(*
	Owned collection of OTLP key-value attributes used across telemetry domains.
*)
{attribute 'enable_dynamic_creation'}
FUNCTION_BLOCK FB_Attributes
VAR
	_head: POINTER TO ST_LinkedListNode;
	_tail: POINTER TO ST_LinkedListNode;
	_cursor: POINTER TO ST_LinkedListNode;
END_VAR
VAR_OUTPUT
	count: UDINT;
	maxCount: UDINT;
	droppedCount: UDINT;
END_VAR

(* The enforced bound: maxCount, held to MAX_LOOP_COUNT so free always reaches the end. *)
METHOD _capacity : UDINT
_capacity := MIN(THIS^.maxCount, TcOtlp_GVL.MAX_LOOP_COUNT);
END_METHOD

(* The node holding the attribute named key, or 0 when there is none. Does not move the next cursor. *)
METHOD _findNode : POINTER TO ST_LinkedListNode
VAR_INPUT
	key: T_MaxString;
END_VAR
VAR
	_idx: UDINT;
	_node: POINTER TO ST_LinkedListNode;
	_pKv: POINTER TO FB_KeyValue;
END_VAR
_findNode := 0;

_node := THIS^._head;
FOR _idx := 0 TO TcOtlp_GVL.MAX_LOOP_COUNT DO
	IF _node = 0 THEN
		RETURN;
	END_IF
	_pKv := _node^.val;
	IF _pKv <> 0 AND_THEN _pKv^.pKey <> 0 AND_THEN _pKv^.pKey^ = key THEN
		_findNode := _node;
		RETURN;
	END_IF
	_node := _node^.nxt;
END_FOR
END_METHOD

METHOD _mapValueFactoryFailure : E_AttributesFailureReason
VAR_INPUT
	failureReason: E_ValueFactoryFailureReason;
END_VAR
CASE failureReason OF
	E_ValueFactoryFailureReason.SOURCE_POINTER_NULL:
		_mapValueFactoryFailure := E_AttributesFailureReason.KV_VALUE_POINTER_NULL;
	E_ValueFactoryFailureReason.KEY_POINTER_NULL:
		_mapValueFactoryFailure := E_AttributesFailureReason.KV_KEY_POINTER_NULL;
	E_ValueFactoryFailureReason.VALUE_POINTER_NULL:
		_mapValueFactoryFailure := E_AttributesFailureReason.KV_VALUE_POINTER_NULL;
	E_ValueFactoryFailureReason.UNSUPPORTED_VALUE_TYPE:
		_mapValueFactoryFailure := E_AttributesFailureReason.KV_VALUE_TYPE_UNSUPPORTED;
	E_ValueFactoryFailureReason.MEMORY_ALLOCATION_FAILURE:
		_mapValueFactoryFailure := E_AttributesFailureReason.MEMORY_ALLOCATION_FAILURE;
	ELSE
		_mapValueFactoryFailure := E_AttributesFailureReason.KV_VALUE_INVALID;
END_CASE
END_METHOD

(*
	Adds a copy of src's attribute named key, stored under destKey, or under key when destKey is
	empty. An attribute already held under that name is replaced, as with setAttribute. src is
	left unchanged and may be this collection, so an attribute can be copied to a new name in place.
*)
METHOD copyAttribute : BOOL
VAR_IN_OUT
	src: FB_Attributes;
END_VAR
VAR_INPUT
	key: T_MaxString;
	destKey: T_MaxString := '';
END_VAR
VAR_OUTPUT
	failureReason: E_AttributesFailureReason;
END_VAR
VAR
	_pSrc: POINTER TO FB_KeyValue;
	_pDest: POINTER TO FB_KeyValue;
	_factoryFailureReason: E_ValueFactoryFailureReason;
END_VAR
copyAttribute := FALSE;
failureReason := E_AttributesFailureReason.NA;

_pSrc := src.getAttribute(key);
IF _pSrc = 0 THEN
	failureReason := E_AttributesFailureReason.KEY_NOT_FOUND;
	RETURN;
END_IF

IF destKey = '' THEN
	destKey := key;
END_IF

IF NOT ValueFactory.createKeyValue(
	pDest:=_pDest,
	pKey:=ADR(destKey),
	pVal:=_pSrc^.pVal,
	failureReason=>_factoryFailureReason
) THEN
	failureReason := THIS^._mapValueFactoryFailure(_factoryFailureReason);
	RETURN;
END_IF

copyAttribute := THIS^.setAttribute(pValue:=_pDest, failureReason=>failureReason);
// setAttribute only takes ownership on success; release a rejected value
IF _pDest <> 0 THEN
	_pDest^.delete(pSelf:=_pDest);
END_IF
END_METHOD

(*
	Adds a copy of every attribute in src, and carries src's droppedCount over, so the copy
	reports the same loss as the original.
*)
METHOD copyFrom : BOOL
VAR_IN_OUT
	src: FB_Attributes;
END_VAR
VAR_OUTPUT
	failureReason: E_AttributesFailureReason;
END_VAR
VAR
	_idx: UDINT;
	_pSrc: POINTER TO FB_KeyValue;
	_pDest: POINTER TO FB_KeyValue;
	_factoryFailureReason: E_ValueFactoryFailureReason;
END_VAR
copyFrom := FALSE;
failureReason := E_AttributesFailureReason.NA;

THIS^.droppedCount := THIS^.droppedCount + src.droppedCount;
src.reset();
FOR _idx := 0 TO TcOtlp_GVL.MAX_LOOP_COUNT DO
	_pSrc := src.next();
	IF _pSrc = 0 THEN
		copyFrom := failureReason = E_AttributesFailureReason.NA;
		RETURN;
	END_IF
	IF NOT ValueFactory.cloneKeyValue(pDest:=_pDest, pSrc:=_pSrc, failureReason=>_factoryFailureReason) THEN
		failureReason := THIS^._mapValueFactoryFailure(_factoryFailureReason);
		RETURN;
	END_IF
	IF NOT THIS^.setAttribute(pValue:=_pDest, failureReason=>failureReason) THEN
		IF _pDest <> 0 THEN
			_pDest^.delete(pSelf:=_pDest);
		END_IF
		RETURN;
	END_IF
END_FOR

copyFrom := failureReason = E_AttributesFailureReason.NA;
END_METHOD

METHOD FB_Exit : BOOL
VAR_INPUT
	bInCopyCode: BOOL;
END_VAR
IF NOT bInCopyCode THEN
	THIS^.free();
END_IF
END_METHOD

//FB_Init is always available implicitly and it is used primarily for initialization.
//The return value is not evaluated. For a specific influence, you can also declare the
//methods explicitly and provide additional code there with the standard initialization
//code. You can evaluate the return value.
METHOD FB_Init: BOOL
VAR_INPUT
    bInitRetains: BOOL; // TRUE: the retain variables are initialized (reset warm / reset cold)
    bInCopyCode: BOOL;  // TRUE: the instance will be copied to the copy code afterward (online change) 
	maxCount: UDINT := 20;  
END_VAR
THIS^.maxCount := maxCount;
END_METHOD

(*
	Releases every owned attribute. setAttribute holds count to MAX_LOOP_COUNT, so the loop
	always reaches the end, even if maxCount is lowered after attributes were added. If it ever
	stops early, the unreleased nodes stay in the collection and free returns FALSE, so a later
	call can finish the job.
*)
METHOD free : BOOL
VAR
	_idx: UDINT;
	_node: POINTER TO ST_LinkedListNode;
	_kv: POINTER TO FB_KeyValue;
END_VAR
FOR _idx := 0 TO TcOtlp_GVL.MAX_LOOP_COUNT DO
	IF THIS^._head = 0 THEN
		EXIT;
	END_IF

	_node := THIS^._head;
	THIS^._head := _node^.nxt;
	IF _node^.val <> 0 THEN
		_kv := _node^.val;
		_node^.val := 0;
		_kv^.delete(pSelf:=_kv);
	END_IF
	__DELETE(_node);
	_node := 0;
	IF THIS^.count > 0 THEN
		THIS^.count := THIS^.count - 1;
	END_IF
END_FOR

IF THIS^._head = 0 THEN
	THIS^._tail := 0;
	THIS^.count := 0;
END_IF
THIS^._cursor := THIS^._head;
free := THIS^._head = 0;
END_METHOD

(*
	Returns the attribute named key, or 0 when there is none. The collection keeps ownership: the
	pointer is borrowed and stays valid only until that attribute is replaced or the collection is
	freed. Does not move the next cursor.
*)
METHOD getAttribute : POINTER TO FB_KeyValue
VAR_INPUT
	key: T_MaxString;
END_VAR
VAR
	_node: POINTER TO ST_LinkedListNode;
END_VAR
getAttribute := 0;

_node := THIS^._findNode(key);
IF _node <> 0 THEN
	getAttribute := _node^.val;
END_IF
END_METHOD

METHOD next : POINTER TO FB_KeyValue
next := 0;

IF THIS^._cursor <> 0 THEN
	next := THIS^._cursor^.val;
	THIS^._cursor := THIS^._cursor^.nxt;
END_IF
END_METHOD

METHOD reset
THIS^._cursor := THIS^._head;
END_METHOD

METHOD setAttribute : BOOL
VAR_IN_OUT
	pValue: POINTER TO FB_KeyValue;
END_VAR
VAR_OUTPUT
	failureReason: E_AttributesFailureReason;
END_VAR
VAR
	_node: POINTER TO ST_LinkedListNode;
	_pVal: POINTER TO FB_KeyValue;
END_VAR
setAttribute := FALSE;
failureReason := E_AttributesFailureReason.NA;

IF pValue = 0 THEN
	failureReason := E_AttributesFailureReason.KV_POINTER_NULL;
	RETURN;
END_IF

IF pValue^.pKey = 0 THEN
	failureReason := E_AttributesFailureReason.KV_KEY_POINTER_NULL;
	RETURN;
END_IF

IF pValue^.pVal = 0 THEN
	failureReason := E_AttributesFailureReason.KV_VALUE_POINTER_NULL;
	RETURN;
END_IF

// replace the value if the key already exists
_node := THIS^._findNode(pValue^.pKey^);
IF _node <> 0 THEN
	_pVal := _node^.val;
	_pVal^.delete(pSelf:=_pVal);
	_node^.val := pValue;
	setAttribute := failureReason = E_AttributesFailureReason.NA;
	pValue := 0;
	RETURN;
END_IF

IF THIS^.count >= THIS^._capacity() THEN
	failureReason := E_AttributesFailureReason.ATTRIBUTE_COUNT_LIMIT_REACHED;
	THIS^.droppedCount := THIS^.droppedCount + 1;
	RETURN;
END_IF

// if it doesn't exist append the key-value pair
_node := __NEW(ST_LinkedListNode);
IF _node = 0 THEN
	failureReason := E_AttributesFailureReason.MEMORY_ALLOCATION_FAILURE;
	RETURN;
END_IF

_node^.val := pValue;
_node^.nxt := 0;

IF THIS^._tail = 0 THEN
	THIS^._head := _node;
	THIS^._cursor := _node;
ELSE
	THIS^._tail^.nxt := _node;
END_IF

THIS^._tail := _node;
THIS^.count := THIS^.count + 1;

// Ownership transfers only after the value has been linked successfully.
pValue := 0;
setAttribute := failureReason = E_AttributesFailureReason.NA;
END_METHOD

METHOD setNumberAttribute : BOOL
VAR_INPUT
	key: T_MaxString;
	value: ANY_NUM;
END_VAR
VAR_OUTPUT
	failureReason: E_AttributesFailureReason;
END_VAR
VAR
	_pKv: POINTER TO FB_KeyValue;
	_pNum: POINTER TO FB_Number;
	_factoryFailureReason: E_ValueFactoryFailureReason;
END_VAR
setNumberAttribute := FALSE;
failureReason := E_AttributesFailureReason.NA;

IF NOT ValueFactory.createNumber_AnyType(
	pDest:=_pNum,
	value:=value,
	failureReason=>_factoryFailureReason
) THEN
	failureReason := THIS^._mapValueFactoryFailure(_factoryFailureReason);
	RETURN;
END_IF

IF NOT ValueFactory.createKeyValue(
	pDest:=_pKv,
	pKey:=ADR(key),
	pVal:=_pNum,
	failureReason=>_factoryFailureReason
) THEN
	failureReason := THIS^._mapValueFactoryFailure(_factoryFailureReason);
	_pNum^.delete(pSelf:=_pNum);
	RETURN;
END_IF
_pNum^.delete(pSelf:=_pNum);  // clean up the _pNum as its cloned in createKeyValue

setNumberAttribute := THIS^.setAttribute(pValue:=_pKv, failureReason=>failureReason);
// setAttribute only takes ownership on success; release a rejected value
IF _pKv <> 0 THEN
	_pKv^.delete(pSelf:=_pKv);
END_IF
END_METHOD

METHOD setNumberAttribute_AnyType : BOOL
VAR_INPUT
	key: T_MaxString;
	value: AnyType;
END_VAR
VAR_OUTPUT
	failureReason: E_AttributesFailureReason;
END_VAR
VAR
	_pKv: POINTER TO FB_KeyValue;
	_pNum: POINTER TO FB_Number;
	_factoryFailureReason: E_ValueFactoryFailureReason;
END_VAR
setNumberAttribute_AnyType := FALSE;
failureReason := E_AttributesFailureReason.NA;

IF NOT ValueFactory.createNumber_AnyType(
	pDest:=_pNum,
	value:=value,
	failureReason=>_factoryFailureReason
) THEN
	failureReason := THIS^._mapValueFactoryFailure(_factoryFailureReason);
	RETURN;
END_IF

IF NOT ValueFactory.createKeyValue(
	pDest:=_pKv,
	pKey:=ADR(key),
	pVal:=_pNum,
	failureReason=>_factoryFailureReason
) THEN
	failureReason := THIS^._mapValueFactoryFailure(_factoryFailureReason);
	_pNum^.delete(pSelf:=_pNum);
	RETURN;
END_IF
_pNum^.delete(pSelf:=_pNum);  // clean up the _pNum as its cloned in createKeyValue

setNumberAttribute_AnyType := THIS^.setAttribute(pValue:=_pKv, failureReason=>failureReason);
// setAttribute only takes ownership on success; release a rejected value
IF _pKv <> 0 THEN
	_pKv^.delete(pSelf:=_pKv);
END_IF
END_METHOD

METHOD setStringAttribute : BOOL
VAR_INPUT
	key: T_MaxString;
	value: T_MaxString;
END_VAR
VAR_OUTPUT
	failureReason: E_AttributesFailureReason;
END_VAR
VAR
	_pKv: POINTER TO FB_KeyValue;
	_pStr: POINTER TO FB_String;
	_factoryFailureReason: E_ValueFactoryFailureReason;
END_VAR
setStringAttribute := FALSE;
failureReason := E_AttributesFailureReason.NA;

IF NOT ValueFactory.createString(
	pDest:=_pStr,
	pString:=ADR(value),
	failureReason=>_factoryFailureReason
) THEN
	failureReason := THIS^._mapValueFactoryFailure(_factoryFailureReason);
	RETURN;
END_IF

IF NOT ValueFactory.createKeyValue(
	pDest:=_pKv,
	pKey:=ADR(key),
	pVal:=_pStr,
	failureReason=>_factoryFailureReason
) THEN
	failureReason := THIS^._mapValueFactoryFailure(_factoryFailureReason);
	_pStr^.delete(pSelf:=_pStr);
	RETURN;
END_IF
_pStr^.delete(pSelf:=_pStr);  // clean up the _pStr as its cloned in createKeyValue

setStringAttribute := THIS^.setAttribute(pValue:=_pKv, failureReason=>failureReason);
// setAttribute only takes ownership on success; release a rejected value
IF _pKv <> 0 THEN
	_pKv^.delete(pSelf:=_pKv);
END_IF
END_METHOD

END_FUNCTION_BLOCK

(* stored: Version 1.1.0.1
   POU FB_Attributes: Id {cf073bde-f48d-4029-b947-e958e98bbb16}, SpecialFunc None
   Method _capacity: Id {5d7c2e1a-8b43-4f6e-9a1d-3c2b7e9f0a64}
   Method _findNode: Id {8e2f6b14-7c39-4d0a-b5e1-94a3c7d2f058}
   Method _mapValueFactoryFailure: Id {b07c94f0-2f89-4b83-a86c-5297aea8b765}
   Method copyAttribute: Id {b754f058-69f8-4057-bad5-234822fe208a}
   Method copyFrom: Id {12dc0284-c0fc-445c-a394-015d07f02ff7}
   Method FB_Exit: Id {686344bf-91ee-4a2a-b059-004362cdb29b}
   Method FB_Init: Id {37f12a41-417f-40ad-87ed-c4eb97312d76}
   Method free: Id {cac7191c-0f7c-4339-b12b-895becc570f8}
   Method getAttribute: Id {51bb0bec-2ec7-474d-bc68-bfc0daab6de0}
   Method next: Id {a8ca5105-d23e-40b3-adba-9bbe23230589}
   Method reset: Id {8ff040db-0c4f-4ccd-95b1-134233b77487}
   Method setAttribute: Id {29d543f3-3e33-4876-b1bf-4a2f0254ef43}
   Method setNumberAttribute: Id {5ce7a6f9-75cf-4bf9-8ec2-655b0a7ea8b4}
   Method setNumberAttribute_AnyType: Id {a633e97e-967c-40bb-9f1d-14d8e2ed4da3}
   Method setStringAttribute: Id {807c259f-0345-4462-a6a8-1359a14a613b} *)
